{region 'Documentation'}
(*!
<summary>Checks that the selected WORD bit differs from the expected Boolean value.</summary>
*)
{endregion}
FUNCTION_BLOCK AssertNotEqualBit_Word EXTENDS AssertionBase
VAR_INPUT
    IN : WORD; //! Actual bitfield.
    BitIndex : USINT; //! Zero-based bit index (0..15); an invalid index produces Error during evaluation.
    Expected : BOOL; //! Forbidden selected bit value.
END_VAR

SUPER^();

{region 'Documentation'}
(*!
<summary>Validates the index before evaluating the selected bit.</summary>
*)
{endregion}
METHOD PROTECTED Assert
VAR
    Mask : WORD;
    ActualBit : BOOL;
    Message : STRING(GVL_Constants.MessageLength);
    ActualText : STRING(GVL_Constants.AssertionValueLength);
END_VAR
VAR CONSTANT
    MaxBitIndex : USINT := 15;
    SingleBitMask : WORD := 16#01;
    NoBitMask : WORD := 16#00;
    HexDigitCount : USINT := 4;
END_VAR
IF NOT EvaluationActive THEN
    RETURN;
END_IF;

IF Result = E_Result.Error THEN
    RETURN;
END_IF;

IF BitIndex > MaxBitIndex THEN
    Message := CONCAT('Assertion error: bit index is outside valid range. BitIndex = ',
        USINT_TO_STRING(BitIndex));
    Message := CONCAT(Message, ', MaxBitIndex = ');
    Message := CONCAT(Message, USINT_TO_STRING(MaxBitIndex));
    Message := CONCAT(Message, '.');
    Error(Message := Message);
    RETURN;
END_IF;

IF Result = E_Result.Failed THEN
    RETURN;
END_IF;

Mask := SHL(SingleBitMask, BitIndex);
ActualBit := (IN AND Mask) <> NoBitMask;

IF ActualBit = Expected THEN
    ActualText := CreateAssertionTextValue_Hex(Value := WORD_TO_LWORD(IN),
        DigitCount := HexDigitCount);
    Message := CONCAT('Assertion failed: bit value matches forbidden value. BitIndex = ',
        USINT_TO_STRING(BitIndex));
    Message := CONCAT(Message, ', NotExpected = ');
    Message := CONCAT(Message, BOOL_TO_STRING(Expected));
    Message := CONCAT(Message, ', Actual = ');
    Message := CONCAT(Message, BOOL_TO_STRING(ActualBit));
    Message := CONCAT(Message, ', Value = ');
    Message := CONCAT(Message, ActualText);
    Message := CONCAT(Message, '.');
    Fail(Message := Message);
    RETURN;
END_IF;

Pass();
END_METHOD

END_FUNCTION_BLOCK

(* stored: Version 1.1.0.1
   POU AssertNotEqualBit_Word: Id {7e18ff8c-d4b6-49be-bd8d-a1eae24b75d8}, SpecialFunc None
   Folder Internal: Id {ed5990a1-d93f-4678-912b-5fc6500384ea}
   Method Assert: Id {edfae680-a186-4159-a6c7-24bebdc0e221} *)
